Staubli VAL3: frameItem.pjx

--- frameItem.pjx ---
Parameters version=s8.10.3Cs9_BS2093 stackSize=5000 millimeterUnit=true
Program file=start.pgx
Program file=stop.pgx
Data file=frameItem.dtx

--- frameItem.dtx ---
public string sName
public frame fFrame = {fatherId=world[0]}
public pointRx pPointRx[3]
  [0] = {fatherId=world[0]}
  [1] = {fatherId=world[0]}
  [2] = {fatherId=world[0]}

--- start.pgx ---
program start()
begin
end

--- stop.pgx ---
program stop()
begin
end
